(* IEC 61131-3 sources: sis-interlock-demo/src/POUs/Sis/F_SisCrc16Byte, 2 files *)

(* ---- F_SisCrc16Byte.decl.st ---- *)
// Назначение: шаг CRC-16/CCITT-FALSE по одному байту: полином 16#1021, без отражения, старший
//             бит первым (раздел 6.8).
// Автор:      kr0nsch
// Версия:     0.1.0
// Документ:   docs/DESIGN.md, раздел «6.8 Конфигурация и CRC»
// ВНИМАНИЕ:   код демонстрационный и не предназначен для систем безопасности. Реальная ПАЗ
//             требует определения SIL, сертифицированных аппаратных и программных средств
//             и валидации по ГОСТ Р МЭК 61511.
FUNCTION F_SisCrc16Byte : WORD
VAR_INPUT
    wCrc  : WORD;    // CRC до этого байта
    bData : BYTE;    // очередной байт
END_VAR
VAR
    wReg  : WORD;    // регистр CRC
    uiBit : UINT;    // номер шага по битам
END_VAR

(* ---- F_SisCrc16Byte.impl.st ---- *)
wReg := wCrc XOR SHL(BYTE_TO_WORD(bData), GVL_Const.BITS_PER_BYTE);
FOR uiBit := 1 TO GVL_Const.BITS_PER_BYTE DO
    IF (wReg AND GVL_Const.CRC16_MSB) <> 0 THEN
        wReg := SHL(wReg, 1) XOR GVL_Const.CRC16_POLY;
    ELSE
        wReg := SHL(wReg, 1);
    END_IF
END_FOR
F_SisCrc16Byte := wReg;
